Universal Robots URScript: letra_D.script

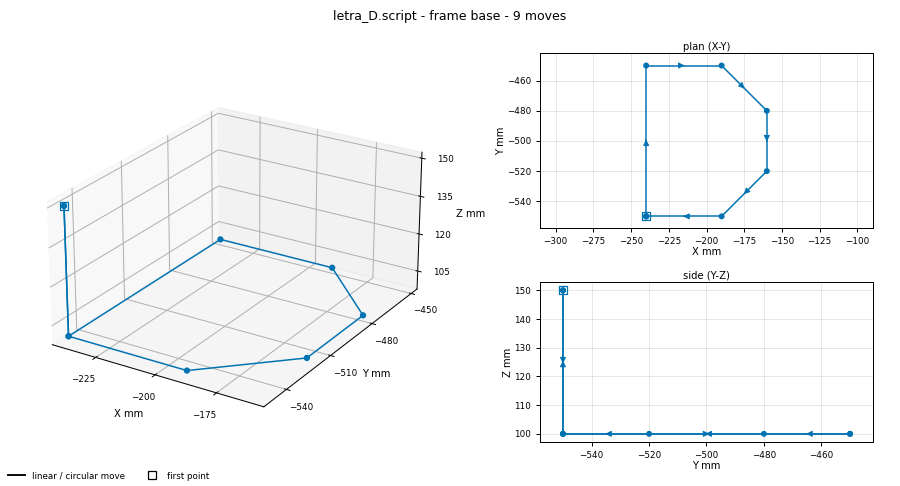
[picture p0: tool path of letra_D.script in frame base, 9 of 9 moves have a stored position in this frame; points joined in program order, loops and branches not executed]
# Letra D - Daniel
movel(p[-0.240, -0.550, 0.150, 3.1416, 0, 0], a=0.5, v=0.1)
movel(p[-0.240, -0.550, 0.100, 3.1416, 0, 0], a=0.5, v=0.1)
movel(p[-0.240, -0.450, 0.100, 3.1416, 0, 0], a=0.5, v=0.1)
movel(p[-0.190, -0.450, 0.100, 3.1416, 0, 0], a=0.5, v=0.1)
movel(p[-0.160, -0.480, 0.100, 3.1416, 0, 0], a=0.5, v=0.1)
movel(p[-0.160, -0.520, 0.100, 3.1416, 0, 0], a=0.5, v=0.1)
movel(p[-0.190, -0.550, 0.100, 3.1416, 0, 0], a=0.5, v=0.1)
movel(p[-0.240, -0.550, 0.100, 3.1416, 0, 0], a=0.5, v=0.1)
movel(p[-0.240, -0.550, 0.150, 3.1416, 0, 0], a=0.5, v=0.1)
